(* IEC 61131-3 sources: volt/packages/volt-lsp-iec/test-corpus/pro2193/Device/Plc Logic/Application/09 Misc/Library Manager/SysSocket Implementation, 44 files *)

(* ---- SYSSOCKACCEPT.pou ---- *)
FUNCTION SYSSOCKACCEPT : RTS_IEC_HANDLE
VAR_INPUT
	HSOCKET : RTS_IEC_HANDLE;
	PSOCKADDR : POINTER TO SOCKADDRESS;
	PDISOCKADDRSIZE : POINTER TO DINT;
	PRESULT : POINTER TO RTS_IEC_RESULT;
END_VAR
END_FUNCTION

(* ---- SYSSOCKBIND.pou ---- *)
FUNCTION SYSSOCKBIND : RTS_IEC_RESULT
VAR_INPUT
	HSOCKET : RTS_IEC_HANDLE;
	PSOCKADDR : POINTER TO SOCKADDRESS;
	DISOCKADDRSIZE : DINT;
END_VAR
END_FUNCTION

(* ---- SYSSOCKCLOSE.pou ---- *)
FUNCTION SYSSOCKCLOSE : RTS_IEC_RESULT
VAR_INPUT
	HSOCKET : RTS_IEC_HANDLE;
END_VAR
END_FUNCTION

(* ---- SYSSOCKCLOSEUDP.pou ---- *)
FUNCTION SYSSOCKCLOSEUDP : RTS_IEC_RESULT
VAR_INPUT
	HSOCKETUDP : RTS_IEC_HANDLE;
END_VAR
END_FUNCTION

(* ---- SYSSOCKCONNECT.pou ---- *)
FUNCTION SYSSOCKCONNECT : RTS_IEC_RESULT
VAR_INPUT
	HSOCKET : RTS_IEC_HANDLE;
	PSOCKADDR : POINTER TO SOCKADDRESS;
	DISOCKADDRSIZE : DINT;
END_VAR
END_FUNCTION

(* ---- SYSSOCKCREATE.pou ---- *)
FUNCTION SYSSOCKCREATE : RTS_IEC_HANDLE
VAR_INPUT
	IADDRESSFAMILY : INT;
	DITYPE : DINT;
	DIPROTOCOL : DINT;
	PRESULT : POINTER TO RTS_IEC_RESULT;
END_VAR
END_FUNCTION

(* ---- SYSSOCKCREATEUDP.pou ---- *)
FUNCTION SYSSOCKCREATEUDP : RTS_IEC_HANDLE
VAR_INPUT
	DISENDPORT : DINT;
	DIRECVPORT : DINT;
	PRESULT : POINTER TO RTS_IEC_RESULT;
END_VAR
END_FUNCTION

(* ---- SYSSOCKFDINIT.pou ---- *)
FUNCTION SYSSOCKFDINIT : RTS_IEC_RESULT
VAR_INPUT
	HSOCKET : RTS_IEC_HANDLE;
	PFS : REFERENCE TO SOCKET_FD_SET;
END_VAR
END_FUNCTION

(* ---- SYSSOCKFDISSET.pou ---- *)
FUNCTION SYSSOCKFDISSET : BOOL
VAR_INPUT
	HSOCKET : RTS_IEC_HANDLE;
	PFS : REFERENCE TO SOCKET_FD_SET;
END_VAR
END_FUNCTION

(* ---- SYSSOCKFDZERO.pou ---- *)
FUNCTION SYSSOCKFDZERO : RTS_IEC_RESULT
VAR_INPUT
	PFS : REFERENCE TO SOCKET_FD_SET;
END_VAR
END_FUNCTION

(* ---- SYSSOCKGETFIRSTADAPTERINFO.pou ---- *)
FUNCTION SYSSOCKGETFIRSTADAPTERINFO : RTS_IEC_HANDLE
VAR_INPUT
	PADAPTERINFO : POINTER TO SOCK_ADAPTER_INFORMATION;
	PUXIADAPTERINFOSIZE : POINTER TO __UXINT;
	PRESULT : POINTER TO RTS_IEC_RESULT;
END_VAR
END_FUNCTION

(* ---- SYSSOCKGETHOSTBYNAME.pou ---- *)
FUNCTION SYSSOCKGETHOSTBYNAME : RTS_IEC_RESULT
VAR_INPUT
	SZHOSTNAME : REFERENCE TO STRING;
	PHOST : POINTER TO SOCK_HOSTENT;
END_VAR
END_FUNCTION

(* ---- SYSSOCKGETHOSTNAME.pou ---- *)
FUNCTION SYSSOCKGETHOSTNAME : RTS_IEC_RESULT
VAR_INPUT
	SZHOSTNAME : REFERENCE TO STRING;
	DINAMELEN : DINT;
END_VAR
END_FUNCTION

(* ---- SYSSOCKGETNEXTADAPTERINFO.pou ---- *)
FUNCTION SYSSOCKGETNEXTADAPTERINFO : RTS_IEC_HANDLE
VAR_INPUT
	HPREVADAPTER : RTS_IEC_HANDLE;
	PADAPTERINFO : POINTER TO SOCK_ADAPTER_INFORMATION;
	PUXIADAPTERINFOSIZE : POINTER TO __UXINT;
	PRESULT : POINTER TO RTS_IEC_RESULT;
END_VAR
END_FUNCTION

(* ---- SYSSOCKGETOPTION.pou ---- *)
FUNCTION SYSSOCKGETOPTION : RTS_IEC_RESULT
VAR_INPUT
	HSOCKET : RTS_IEC_HANDLE;
	DILEVEL : DINT;
	DIOPTION : DINT;
	PDIOPTIONVALUE : POINTER TO DINT;
	PDIOPTIONLEN : POINTER TO DINT;
END_VAR
END_FUNCTION

(* ---- SYSSOCKGETOSHANDLE.pou ---- *)
FUNCTION SYSSOCKGETOSHANDLE : RTS_IEC_HANDLE
VAR_INPUT
	HSOCKETUDP : RTS_IEC_HANDLE;
END_VAR
END_FUNCTION

(* ---- SYSSOCKGETPEERNAME.pou ---- *)
FUNCTION SYSSOCKGETPEERNAME : RTS_IEC_RESULT
VAR_INPUT
	HSOCKET : RTS_IEC_HANDLE;
	PSOCKADDR : POINTER TO SOCKADDRESS;
	PDISOCKADDRSIZE : POINTER TO DINT;
END_VAR
END_FUNCTION

(* ---- SYSSOCKGETRECVSIZEUDP.pou ---- *)
FUNCTION SYSSOCKGETRECVSIZEUDP : __XINT
VAR_INPUT
	HSOCKETUDP : RTS_IEC_HANDLE;
	DITIMEOUT : DINT;
	PRESULT : POINTER TO RTS_IEC_RESULT;
END_VAR
END_FUNCTION

(* ---- SYSSOCKGETSOCKNAME.pou ---- *)
FUNCTION SYSSOCKGETSOCKNAME : RTS_IEC_RESULT
VAR_INPUT
	HSOCKET : RTS_IEC_HANDLE;
	PSOCKADDR : POINTER TO SOCKADDRESS;
	PDISOCKADDRSIZE : POINTER TO DINT;
END_VAR
END_FUNCTION

(* ---- SYSSOCKGETSUBNETMASK.pou ---- *)
FUNCTION SYSSOCKGETSUBNETMASK : RTS_IEC_RESULT
VAR_INPUT
	SZIPADDRESS : REFERENCE TO STRING;
	SZSUBNETMASK : REFERENCE TO STRING;
	DIMAXSUGNETMASK : DINT;
END_VAR
END_FUNCTION

(* ---- SYSSOCKHTONL.pou ---- *)
FUNCTION SYSSOCKHTONL : UDINT
VAR_INPUT
	ULHOST : UDINT;
END_VAR
END_FUNCTION

(* ---- SYSSOCKHTONS.pou ---- *)
FUNCTION SYSSOCKHTONS : WORD
VAR_INPUT
	USHOST : WORD;
END_VAR
END_FUNCTION

(* ---- SYSSOCKINETADDR.pou ---- *)
FUNCTION SYSSOCKINETADDR : RTS_IEC_RESULT
VAR_INPUT
	SZIPADDRESS : REFERENCE TO STRING;
	PINADDR : POINTER TO UDINT;
END_VAR
END_FUNCTION

(* ---- SYSSOCKINETNTOA.pou ---- *)
FUNCTION SYSSOCKINETNTOA : RTS_IEC_RESULT
VAR_INPUT
	PINADDR : POINTER TO INADDR;
	SZIPADDR : REFERENCE TO STRING;
	DIIPADDRSIZE : DINT;
END_VAR
END_FUNCTION

(* ---- SYSSOCKIOCTL.pou ---- *)
FUNCTION SYSSOCKIOCTL : RTS_IEC_RESULT
VAR_INPUT
	HSOCKET : RTS_IEC_HANDLE;
	DICOMMAND : DINT;
	PDIPARAMETER : POINTER TO DINT;
END_VAR
END_FUNCTION

(* ---- SYSSOCKLISTEN.pou ---- *)
FUNCTION SYSSOCKLISTEN : RTS_IEC_RESULT
VAR_INPUT
	HSOCKET : RTS_IEC_HANDLE;
	DIMAXCONNECTIONS : DINT;
END_VAR
END_FUNCTION

(* ---- SYSSOCKNTOHL.pou ---- *)
FUNCTION SYSSOCKNTOHL : UDINT
VAR_INPUT
	ULNET : UDINT;
END_VAR
END_FUNCTION

(* ---- SYSSOCKNTOHS.pou ---- *)
FUNCTION SYSSOCKNTOHS : WORD
VAR_INPUT
	USNET : WORD;
END_VAR
END_FUNCTION

(* ---- SYSSOCKPING.pou ---- *)
FUNCTION SYSSOCKPING : RTS_IEC_RESULT
VAR_INPUT
	SZIPADDRESS : REFERENCE TO STRING;
	ULTIMEOUT : UDINT;
	PULREPLYTIME : POINTER TO UDINT;
END_VAR
END_FUNCTION

(* ---- SYSSOCKRECV.pou ---- *)
FUNCTION SYSSOCKRECV : __XINT
VAR_INPUT
	HSOCKET : RTS_IEC_HANDLE;
	PBYBUFFER : POINTER TO BYTE;
	DIBUFFERSIZE : __XINT;
	DIFLAGS : DINT;
	PRESULT : POINTER TO RTS_IEC_RESULT;
END_VAR
END_FUNCTION

(* ---- SYSSOCKRECVFROM.pou ---- *)
FUNCTION SYSSOCKRECVFROM : __XINT
VAR_INPUT
	HSOCKET : RTS_IEC_HANDLE;
	PBYBUFFER : POINTER TO BYTE;
	DIBUFFERSIZE : __XINT;
	DIFLAGS : DINT;
	PSOCKADDR : POINTER TO SOCKADDRESS;
	DISOCKADDRSIZE : DINT;
	PRESULT : POINTER TO RTS_IEC_RESULT;
END_VAR
END_FUNCTION

(* ---- SYSSOCKRECVFROMUDP.pou ---- *)
FUNCTION SYSSOCKRECVFROMUDP : __XINT
VAR_INPUT
	HSOCKETUDP : RTS_IEC_HANDLE;
	PBYDATA : POINTER TO BYTE;
	DIDATASIZE : __XINT;
	PREPLY : POINTER TO UDP_REPLY;
	PRESULT : POINTER TO RTS_IEC_RESULT;
END_VAR
END_FUNCTION

(* ---- SYSSOCKRECVFROMUDP2.pou ---- *)
FUNCTION SYSSOCKRECVFROMUDP2 : __XINT
VAR_INPUT
	HSOCKETUDP : RTS_IEC_HANDLE;
	PBYDATA : POINTER TO BYTE;
	DIDATASIZE : __XINT;
	PREPLY : POINTER TO UDP_REPLY2;
	PRESULT : POINTER TO RTS_IEC_RESULT;
END_VAR
END_FUNCTION

(* ---- SYSSOCKRECVMSG.pou ---- *)
FUNCTION SYSSOCKRECVMSG : __XINT
VAR_INPUT
	HSOCKET : RTS_IEC_HANDLE;
	PMESSAGE : POINTER TO SOCK_RECVMSG_MSG;
	FLAGS : DWORD;
	PRESULT : POINTER TO RTS_IEC_RESULT;
END_VAR
END_FUNCTION

(* ---- SYSSOCKSELECT.pou ---- *)
FUNCTION SYSSOCKSELECT : RTS_IEC_RESULT
VAR_INPUT
	DIWIDTH : DINT;
	PFDREAD : POINTER TO SOCKET_FD_SET;
	PFDWRITE : POINTER TO SOCKET_FD_SET;
	PFDEXCEPT : POINTER TO SOCKET_FD_SET;
	PTVTIMEOUT : POINTER TO SOCKET_TIMEVAL;
	PDIREADY : POINTER TO DINT;
END_VAR
END_FUNCTION

(* ---- SYSSOCKSEND.pou ---- *)
FUNCTION SYSSOCKSEND : __XINT
VAR_INPUT
	HSOCKET : RTS_IEC_HANDLE;
	PBYBUFFER : POINTER TO BYTE;
	DIBUFFERSIZE : __XINT;
	DIFLAGS : DINT;
	PRESULT : POINTER TO RTS_IEC_RESULT;
END_VAR
END_FUNCTION

(* ---- SYSSOCKSENDTO.pou ---- *)
FUNCTION SYSSOCKSENDTO : __XINT
VAR_INPUT
	HSOCKET : RTS_IEC_HANDLE;
	PBYBUFFER : POINTER TO BYTE;
	DIBUFFERSIZE : __XINT;
	DIFLAGS : DINT;
	PSOCKADDR : POINTER TO SOCKADDRESS;
	DISOCKADDRSIZE : DINT;
	PRESULT : POINTER TO RTS_IEC_RESULT;
END_VAR
END_FUNCTION

(* ---- SYSSOCKSENDTOUDP.pou ---- *)
FUNCTION SYSSOCKSENDTOUDP : __XINT
VAR_INPUT
	HSOCKETUDP : RTS_IEC_HANDLE;
	DIPORT : DINT;
	SZDESTADDRESS : REFERENCE TO STRING;
	PBYDATA : POINTER TO BYTE;
	DIDATASIZE : __XINT;
	PRESULT : POINTER TO RTS_IEC_RESULT;
END_VAR
END_FUNCTION

(* ---- SYSSOCKSETDEFAULTGATEWAY.pou ---- *)
FUNCTION SYSSOCKSETDEFAULTGATEWAY : RTS_IEC_RESULT
VAR_INPUT
	WSADAPTERNAME : REFERENCE TO WSTRING;
	GATEWAYADDR : REFERENCE TO INADDR;
END_VAR
END_FUNCTION

(* ---- SYSSOCKSETIPADDRESS.pou ---- *)
FUNCTION SYSSOCKSETIPADDRESS : RTS_IEC_RESULT
VAR_INPUT
	SZCARD : REFERENCE TO STRING;
	SZIPADDRESS : REFERENCE TO STRING;
END_VAR
END_FUNCTION

(* ---- SYSSOCKSETIPADDRESSANDNETMASK.pou ---- *)
FUNCTION SYSSOCKSETIPADDRESSANDNETMASK : RTS_IEC_RESULT
VAR_INPUT
	WSADAPTERNAME : REFERENCE TO WSTRING;
	IPADDR : REFERENCE TO INADDR;
	NETMASK : REFERENCE TO INADDR;
END_VAR
END_FUNCTION

(* ---- SYSSOCKSETOPTION.pou ---- *)
FUNCTION SYSSOCKSETOPTION : RTS_IEC_RESULT
VAR_INPUT
	HSOCKET : RTS_IEC_HANDLE;
	DILEVEL : DINT;
	DIOPTION : DINT;
	PDIOPTIONVALUE : POINTER TO DINT;
	DIOPTIONLEN : DINT;
END_VAR
END_FUNCTION

(* ---- SYSSOCKSETSUBNETMASK.pou ---- *)
FUNCTION SYSSOCKSETSUBNETMASK : RTS_IEC_RESULT
VAR_INPUT
	SZIPADDRESS : REFERENCE TO STRING;
	SZSUBNETMASK : REFERENCE TO STRING;
END_VAR
END_FUNCTION

(* ---- SYSSOCKSHUTDOWN.pou ---- *)
FUNCTION SYSSOCKSHUTDOWN : RTS_IEC_RESULT
VAR_INPUT
	HSOCKET : RTS_IEC_HANDLE;
	DIHOW : DINT;
END_VAR
END_FUNCTION
